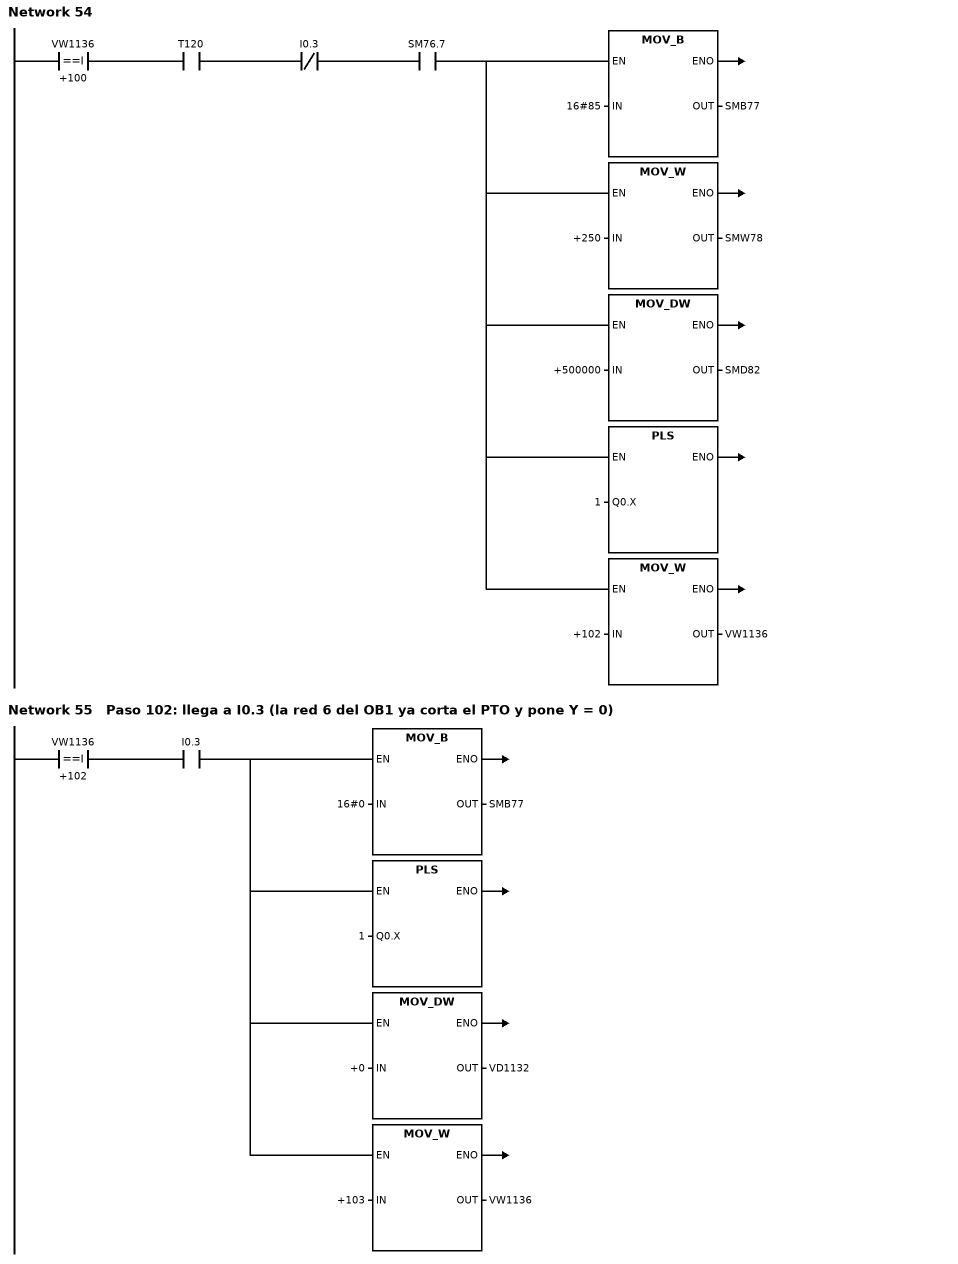
[picture p24: SBR4 networks 54-55]
Network 54
LDW=   VW1136, +100
A      T120
AN     I0.3
A      SM76.7
MOVB   16#85, SMB77
MOVW   +250, SMW78
MOVD   +500000, SMD82
PLS    1
MOVW   +102, VW1136
Network 55 //  Paso 102: llega a I0.3 (la red 6 del OB1 ya corta el PTO y pone Y = 0)
LDW=   VW1136, +102
A      I0.3
MOVB   16#0, SMB77
PLS    1
MOVD   +0, VD1132
MOVW   +103, VW1136
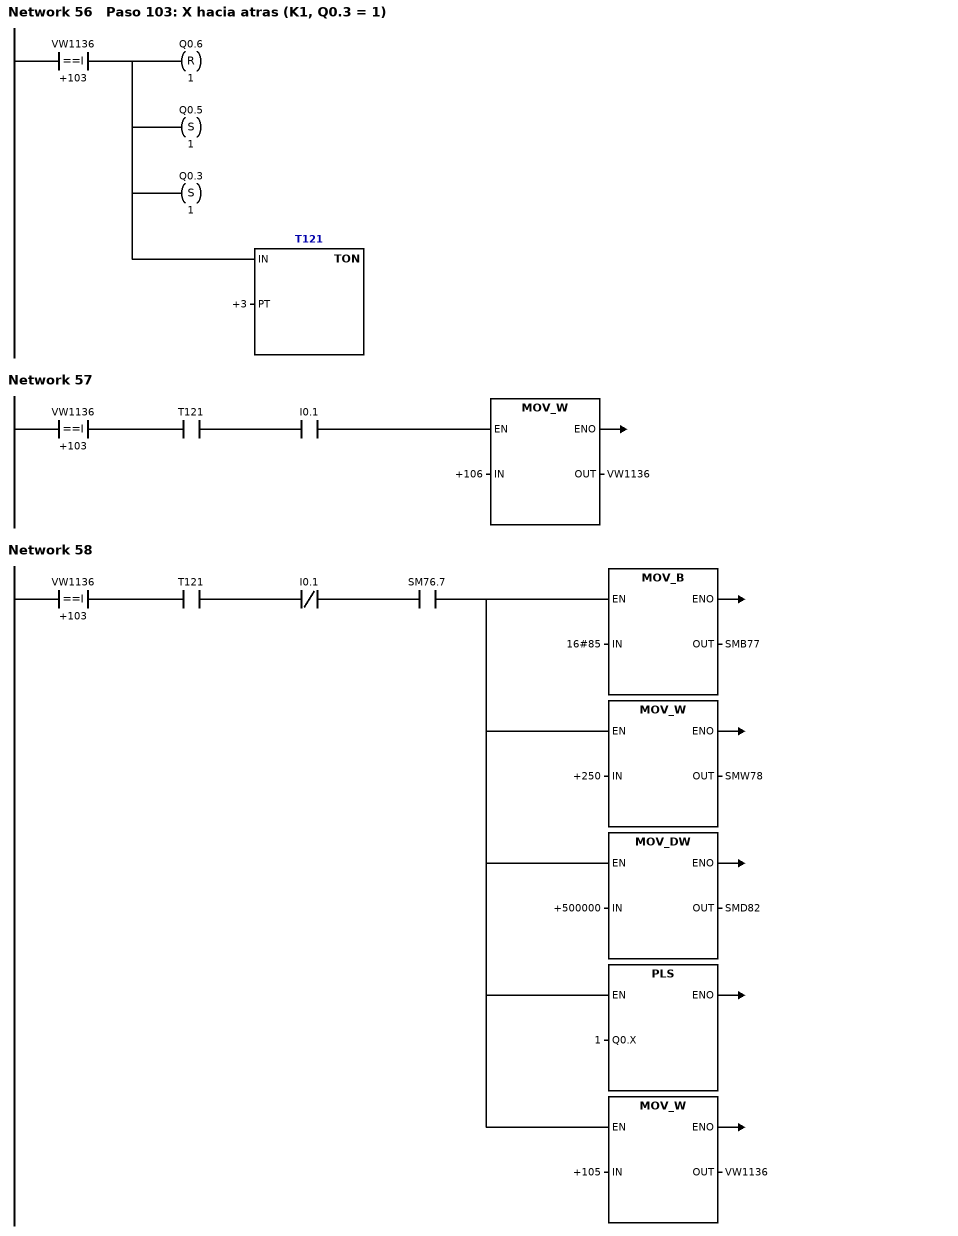
Network 56 //  Paso 103: X hacia atras (K1, Q0.3 = 1)
LDW=   VW1136, +103
R      Q0.6, 1
S      Q0.5, 1
S      Q0.3, 1
TON    T121, +3
Network 57
LDW=   VW1136, +103
A      T121
A      I0.1
MOVW   +106, VW1136
Network 58
LDW=   VW1136, +103
A      T121
AN     I0.1
A      SM76.7
MOVB   16#85, SMB77
MOVW   +250, SMW78
MOVD   +500000, SMD82
PLS    1
MOVW   +105, VW1136
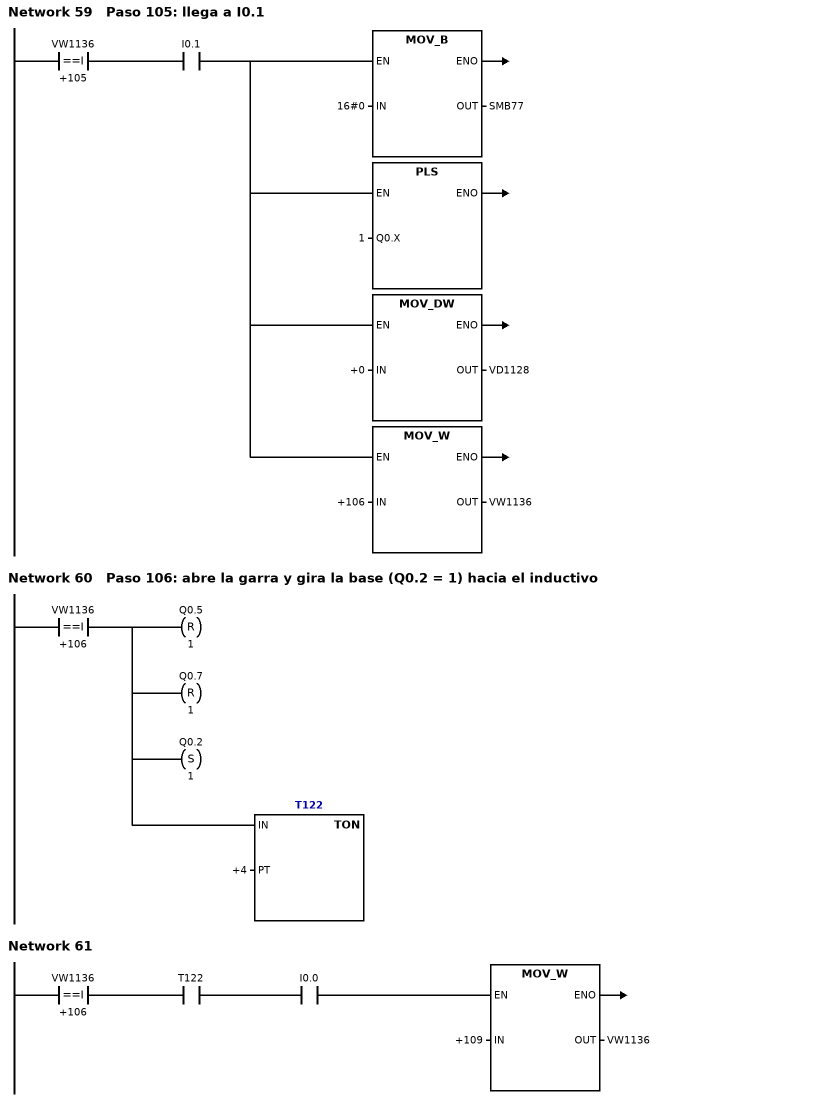
Network 59 //  Paso 105: llega a I0.1
LDW=   VW1136, +105
A      I0.1
MOVB   16#0, SMB77
PLS    1
MOVD   +0, VD1128
MOVW   +106, VW1136
Network 60 //  Paso 106: abre la garra y gira la base (Q0.2 = 1) hacia el inductivo
LDW=   VW1136, +106
R      Q0.5, 1
R      Q0.7, 1
S      Q0.2, 1
TON    T122, +4
Network 61
LDW=   VW1136, +106
A      T122
A      I0.0
MOVW   +109, VW1136
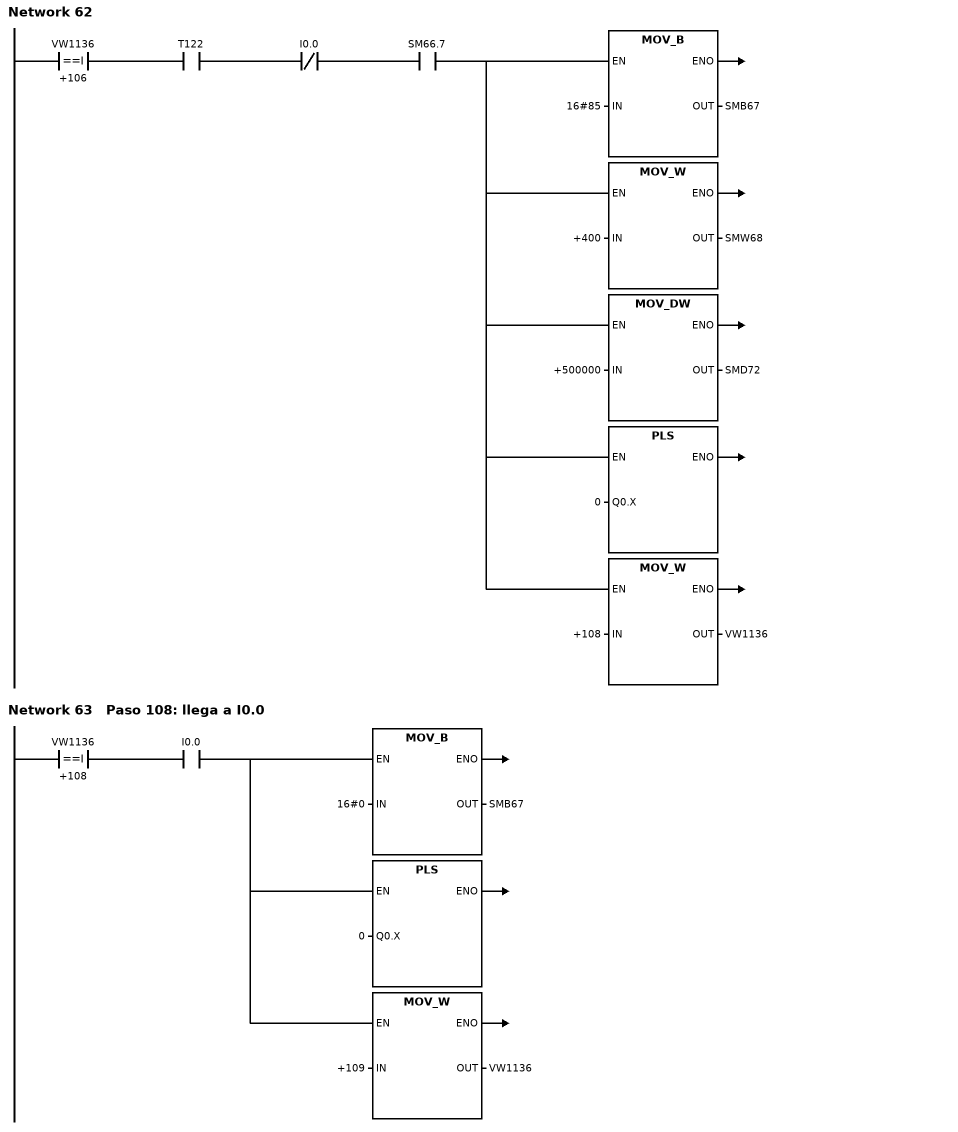
Network 62
LDW=   VW1136, +106
A      T122
AN     I0.0
A      SM66.7
MOVB   16#85, SMB67
MOVW   +400, SMW68
MOVD   +500000, SMD72
PLS    0
MOVW   +108, VW1136
Network 63 //  Paso 108: llega a I0.0
LDW=   VW1136, +108
A      I0.0
MOVB   16#0, SMB67
PLS    0
MOVW   +109, VW1136
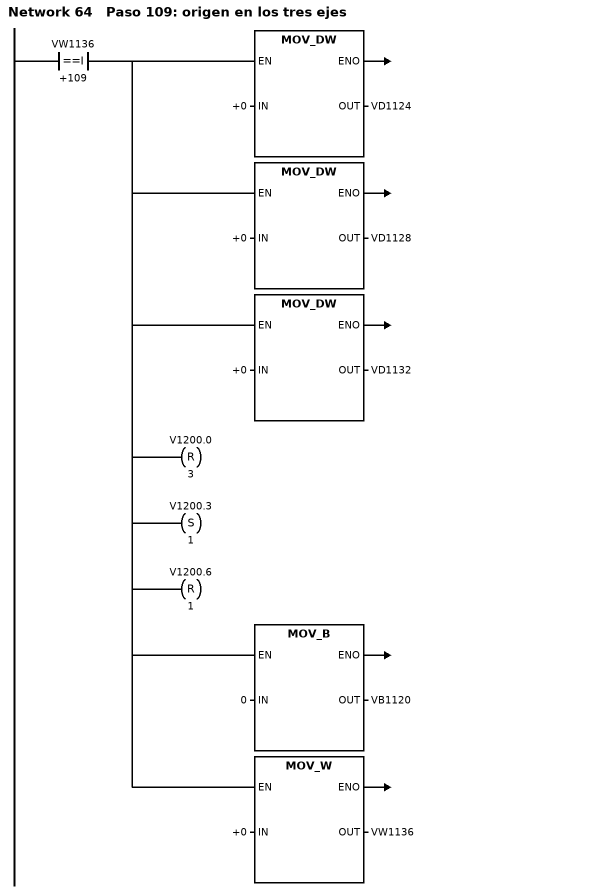
Network 64 //  Paso 109: origen en los tres ejes
LDW=   VW1136, +109
MOVD   +0, VD1124
MOVD   +0, VD1128
MOVD   +0, VD1132
R      V1200.0, 3
S      V1200.3, 1
R      V1200.6, 1
MOVB   0, VB1120
MOVW   +0, VW1136
END_SUBROUTINE_BLOCK
